// TIA Portal V21 export
// export: Created 2000-01-01T00:00:00.0000000Z, ExportSetting None
TYPE "UDT_HMI_FIO_PickAndPlace"
   STRUCT
      bManualMode { ExternalWritable := 'False'} : Bool;   // TRUE: 手动模式, FALSE: 自动模式
      bStartCmd { ExternalWritable := 'False'} : Bool;   // HMI启动触发
      bStopCmd { ExternalWritable := 'False'} : Bool;   // HMI停止触发
      bResetCmd { ExternalWritable := 'False'} : Bool;   // HMI故障复位触发
      bManualMoveX { ExternalWritable := 'False'} : Bool;   // 手动驱动X轴伸出
      bManualMoveZ { ExternalWritable := 'False'} : Bool;   // 手动驱动Z轴下降
      bManualGrab { ExternalWritable := 'False'} : Bool;   // 手动吸盘吸气
      tAxisMoveTime { ExternalWritable := 'False'} : Time;   // 单步气缸动作到位稳定延时（默认 T#600ms）
      tStepTimeout { ExternalWritable := 'False'} : Time;   // 单步动作超时报警时间（默认 T#4s）
      iCurrentStep { ExternalWritable := 'False'} : Int;   // 状态反馈：当前步序
      diPickedCount { ExternalWritable := 'False'} : DInt;   // 状态反馈：累计搬运完成件数
      bRunning { ExternalWritable := 'False'} : Bool;   // 状态反馈：运行中
      bFault { ExternalWritable := 'False'} : Bool;   // 状态反馈：故障标志
      wStatus { ExternalWritable := 'False'} : Word;   // 状态码：16#0000正常, 16#7000待机, 16#8401动作或抓取超时, 16#8402急停切断
   END_STRUCT;
END_TYPE
